(* IEC 61131-3 sources: teller/JD_Teller_LC2_V11/Network/HardwareNet, 1 file *)

(* ---- ONE_HardwareNet_Table.st ---- *)
#define OBJECTS_CONFIG

#include <.\lsl_st_can.h>
#include <.\lsl_st_hardwaretree.h>
//Define part of class HwBaseCDIAS
// Defines for Mutex Generation
#define CDIAS_STR_MUTEX_NAME_SEPERATOR ".."
#define CDIAS_MUTEX_NAME_END_LENGTH 5
#define CDIAS_MUTEX_NAME_MAX_LENGTH 32
//Define part of class CIO0xx
#define ID_CIO0xx 28

#define ID_CIO011 1
#define ID_CIO012 2
#define ID_CIO013 3
#define ID_CIO014 4
#define ID_CIO016 6
#define ID_CIO017 7

#define CIO0xx_Errormask 2#1111111110001111
//Define part of class Varan_Base
#ifndef _T_VARANBASE_H
#define _T_VARANBASE_H

#define	VARAN_PLL_OFFSET		16#0140
#define VARAN_MULTIPLE_OFFSET	16#01AC

// version of serial number validation (16#10 = 1.0)
#define SERNO_VALIDATION_VERSION 16#10

#define IsTransparent_IS_AVAILABLE

// Defines for Mutex Generation
#define VARAN_STR_MUTEX_NAME_SEPERATOR ".."
#define VARAN_MUTEX_NAME_END_LENGTH 5
#define VARAN_MUTEX_NAME_MAX_LENGTH 32

#endif // _T_VARANBASE_H
#include <.\lsl_st_pci.h>
#include "..\..\Class\DiasMasterMain\DiasMasterMain.h"
#include <.\lsl_st_kernel.h>
//Define part of class EEPROM
// Defines for Mutex Geeration
#define EEPROM_STR_MUTEX_NAME_SEPERATOR ".."
#define EEPROM_MUTEX_NAME_END_LENGTH 5
#define EEPROM_MUTEX_NAME_MAX_LENGTH 32
#include "..\..\Class\HwControl\HwControl.h"
//Define part of class SafetyManager
#define LogBufferSize 1000
#include "..\..\Class\SafetyManager\SafetyManager.h"
//Define part of class Varan_Can
#define VARAN_CAN_OS_VERSION	16#1100 + 226
#define CANBUS_INVALID_VALUE	-2147483393			//16#800000FF
//Define part of class VaranManager
#define SIZE_PAYLOAD_FRAME_HEADER_DO      36  // Const because datasize is in the Payload DOs
#define SIZE_PAYLOAD_IRQ_FRAME_HEADER_DO  38  // Const because datasize is in the Payload DOs

#define VM_MAX_POST_INIT_MODULES  1000
#include "..\..\Class\VaranManager\VaranManager.h"

FUNCTION GLOBAL TAB ONE_HardwareNet
-1$UINT, 0$UINT,
0$UINT, 0$UINT,

46$UDINT,
TO_UDINT(529317953), "_CanLib", 1$UINT, 10$UINT, 0$UINT,
TO_UDINT(4078275645), "_SerLib", 1$UINT, 31$UINT, 0$UINT,
TO_UDINT(781409069), "_VaranCanLib", 1$UINT, 10$UINT, 1$UINT,
TO_UDINT(415874427), "_VaranCanLibOS", 1$UINT, 10$UINT, 1$UINT,
TO_UDINT(3827919523), "_VaranSerLibOS", 1$UINT, 20$UINT, 3$UINT,
TO_UDINT(3907636883), "CAICIOAInputChannel", 2$UINT, 20$UINT, 2$UINT,
TO_UDINT(2472734913), "CAIInputChannel", 2$UINT, 20$UINT, 0$UINT,
TO_UDINT(1046309609), "CDias2DataMover", 1$UINT, 50$UINT, 1$UINT,
TO_UDINT(706219532), "ChannelBaseData", 1$UINT, 0$UINT, 0$UINT,
TO_UDINT(3340137983), "ChannelBaseDataWriteOnly", 1$UINT, 0$UINT, 0$UINT,
TO_UDINT(454909577), "CIO011_IM", 2$UINT, 50$UINT, 1$UINT,
TO_UDINT(2636333112), "CIO0xx", 2$UINT, 40$UINT, 0$UINT,
TO_UDINT(3867554050), "CIOOutputChannel", 2$UINT, 20$UINT, 1$UINT,
TO_UDINT(495304727), "CIV521", 1$UINT, 61$UINT, 1$UINT,
TO_UDINT(2756859380), "CIV_Base", 2$UINT, 61$UINT, 0$UINT,
TO_UDINT(658675781), "DAIInputChnl", 2$UINT, 10$UINT, 0$UINT,
TO_UDINT(3820159437), "Dias2DataMover", 1$UINT, 50$UINT, 1$UINT,
TO_UDINT(2647887450), "DiasMaster", 2$UINT, 30$UINT, 0$UINT,
TO_UDINT(3069482179), "DiasMasterC", 1$UINT, 70$UINT, 0$UINT,
TO_UDINT(3792535737), "DiasMasterMain", 2$UINT, 10$UINT, 0$UINT,
TO_UDINT(3076475114), "DiasMasterPostScan", 1$UINT, 0$UINT, 1$UINT,
TO_UDINT(2784851678), "EEPROM", 1$UINT, 11$UINT, 1$UINT,
TO_UDINT(3238133653), "Hub_Base", 1$UINT, 20$UINT, 1$UINT,
TO_UDINT(1770276445), "Hub_Base_Root", 2$UINT, 10$UINT, 1$UINT,
TO_UDINT(1800499398), "HwBaseCDIAS", 2$UINT, 50$UINT, 0$UINT,
TO_UDINT(2471641665), "HwControl", 3$UINT, 0$UINT, 1$UINT,
TO_UDINT(1193052171), "HwControlBase", 1$UINT, 10$UINT, 0$UINT,
TO_UDINT(4260294091), "HWRtPostScan", 1$UINT, 0$UINT, 1$UINT,
TO_UDINT(2326720416), "I2CCDIAS", 1$UINT, 6$UINT, 1$UINT,
TO_UDINT(3953068548), "JD_OR_Teller", 1$UINT, 0$UINT, 1$UINT,
TO_UDINT(2225119864), "MerkerEx", 1$UINT, 18$UINT, 4$UINT,
TO_UDINT(4209775899), "Pulser", 1$UINT, 1$UINT, 1$UINT,
TO_UDINT(3591333481), "RamFile", 1$UINT, 8$UINT, 1$UINT,
TO_UDINT(1799751072), "SafetyManager", 1$UINT, 42$UINT, 1$UINT,
TO_UDINT(1850111279), "String", 1$UINT, 10$UINT, 4$UINT,
TO_UDINT(2898603620), "StringInternal", 1$UINT, 70$UINT, 0$UINT,
TO_UDINT(4187542331), "SyncCall", 1$UINT, 20$UINT, 1$UINT,
TO_UDINT(862125188), "Varan_Base", 2$UINT, 2$UINT, 0$UINT,
TO_UDINT(206510048), "Varan_Can", 1$UINT, 40$UINT, 1$UINT,
TO_UDINT(3752737333), "Varan_DataMover", 1$UINT, 50$UINT, 1$UINT,
TO_UDINT(2940693151), "VaranManager", 2$UINT, 12$UINT, 0$UINT,
TO_UDINT(1989862026), "VaranManager_1", 1$UINT, 43$UINT, 1$UINT,
TO_UDINT(4035182347), "VaranManager_Base", 1$UINT, 20$UINT, 0$UINT,
TO_UDINT(803224590), "VaranManagerPostScan", 1$UINT, 1$UINT, 1$UINT,
TO_UDINT(3232495061), "VirtualBaseInit", 1$UINT, 3$UINT, 0$UINT,
TO_UDINT(1573657038), "WatchdogDias", 2$UINT, 10$UINT, 1$UINT,

1$UINT, TO_UDINT(2726984929), "CIV5211\_VARANCANLIB",

1$UINT, TO_UDINT(3666615371), "CIV5211\_VARANCANLIBOS",

1$UINT, TO_UDINT(2650501396), "CIV5211\_VARANSERLIBOS0",
1$UINT, TO_UDINT(3942400386), "CIV5211\_VARANSERLIBOS1",
1$UINT, TO_UDINT(1945440312), "CIV5211\_VARANSERLIBOS2",

1$UINT, TO_UDINT(3874057698), "CIO011_IM1\CAICIOAINPUTCHANNEL0",
1$UINT, TO_UDINT(2448317812), "CIO011_IM1\CAICIOAINPUTCHANNEL1",

1$UINT, TO_UDINT(407248868), "CIV5211\CDIAS2DATAMOVER",

_NO_ATTR, TO_UDINT(396609901), "CIO011_IM1",

1$UINT, TO_UDINT(325438698), "CIO011_IM1\CIOOUTPUTCHANNEL0",

_NO_ATTR, TO_UDINT(1241008), "CIV5211",

1$UINT, TO_UDINT(569811197), "CIV5211\DIAS2DATAMOVER",

1$UINT, TO_UDINT(2796364169), "CIV5211\DIAS2DATAMOVER\_BASE\DIASMASTERPOSTSCAN",

1$UINT, TO_UDINT(330460277), "CIV5211\DIAS2DATAMOVER\_BASE\EEPROM",

1$UINT, TO_UDINT(2268287070), "CIV5211\HUB_BASE0",

1$UINT, TO_UDINT(1776428101), "VARANMANAGER_11\HUB_BASE_ROOT0",

_NO_ATTR, TO_UDINT(2190789875), "HWCONTROL1",

1$UINT, TO_UDINT(1673205898), "HWCONTROL1\HWRTPOSTSCAN",

1$UINT, TO_UDINT(977257911), "CIV5211\DIAS2DATAMOVER\_BASE\I2CCDIAS",

_NO_ATTR, TO_UDINT(2206833861), "JD_OR1",

1$UINT, TO_UDINT(858933024), "CIO011_IM1\_BASE\_BASE\SERIALNOSTR\MERKEREX0",
1$UINT, TO_UDINT(2644417201), "CIV5211\DIAS2DATAMOVER\_BASE\SYNCCALL\_BASE\SERIALNOSTR\MERKEREX0",
1$UINT, TO_UDINT(3052700284), "CIV5211\DIAS2DATAMOVER\_BASE\WATCHDOGDIAS0\_BASE\SERIALNOSTR\MERKEREX0",
1$UINT, TO_UDINT(2330668179), "CIV5211\_BASE\SERIALNOSTR\MERKEREX0",

_NO_ATTR, TO_UDINT(155437646), "PULSER1",

1$UINT, TO_UDINT(4247336844), "CIV5211\_BASE\SERNOBACKUP",

1$UINT, TO_UDINT(1778590035), "HWCONTROL1\SAFETYMANAGER",

1$UINT, TO_UDINT(2060113651), "CIO011_IM1\_BASE\_BASE\SERIALNOSTR",
1$UINT, TO_UDINT(2623421091), "CIV5211\DIAS2DATAMOVER\_BASE\SYNCCALL\_BASE\SERIALNOSTR",
1$UINT, TO_UDINT(2991369526), "CIV5211\DIAS2DATAMOVER\_BASE\WATCHDOGDIAS0\_BASE\SERIALNOSTR",
1$UINT, TO_UDINT(2961157748), "CIV5211\_BASE\SERIALNOSTR",

1$UINT, TO_UDINT(1225390380), "CIV5211\DIAS2DATAMOVER\_BASE\SYNCCALL",

1$UINT, TO_UDINT(4278451883), "CIV5211\VARAN_CAN",

1$UINT, TO_UDINT(4189409080), "CIV5211\VARAN_DATAMOVER",

_NO_ATTR, TO_UDINT(2395414379), "VARANMANAGER_11",

1$UINT, TO_UDINT(4241828209), "VARANMANAGER_11\_BASE\VARANMASTERPOSTSCAN",

1$UINT, TO_UDINT(2365686840), "CIV5211\DIAS2DATAMOVER\_BASE\WATCHDOGDIAS0",

//Internal connections
0$UDINT,
31$UDINT,
TO_UDINT(8), "SerialNoStr", TO_UDINT(27),
TO_UDINT(8), "CAICIOAInputChannel0", TO_UDINT(5),
TO_UDINT(8), "CAICIOAInputChannel1", TO_UDINT(6),
TO_UDINT(8), "CIOOutputChannel0", TO_UDINT(9),
TO_UDINT(10), "SerialNoStr", TO_UDINT(30),
TO_UDINT(10), "SerNoBackup", TO_UDINT(25),
TO_UDINT(10), "Varan_DataMover", TO_UDINT(33),
TO_UDINT(10), "CDias2DataMover", TO_UDINT(7),
TO_UDINT(10), "Dias2DataMover", TO_UDINT(11),
TO_UDINT(10), "Hub_Base0", TO_UDINT(14),
TO_UDINT(10), "Varan_Can", TO_UDINT(32),
TO_UDINT(10), "_VaranCanLib", TO_UDINT(0),
TO_UDINT(10), "_VaranCanLibOS", TO_UDINT(1),
TO_UDINT(10), "_VaranSerLibOS0", TO_UDINT(2),
TO_UDINT(10), "_VaranSerLibOS1", TO_UDINT(3),
TO_UDINT(10), "_VaranSerLibOS2", TO_UDINT(4),
TO_UDINT(11), "DiasMasterPostScan", TO_UDINT(12),
TO_UDINT(11), "EEPROM", TO_UDINT(13),
TO_UDINT(11), "I2CCDIAS", TO_UDINT(18),
TO_UDINT(11), "WatchdogDias0", TO_UDINT(36),
TO_UDINT(11), "SyncCall", TO_UDINT(31),
TO_UDINT(16), "HWRtPostScan", TO_UDINT(17),
TO_UDINT(16), "SafetyManager", TO_UDINT(26),
TO_UDINT(27), "MerkerEx0", TO_UDINT(20),
TO_UDINT(28), "MerkerEx0", TO_UDINT(21),
TO_UDINT(29), "MerkerEx0", TO_UDINT(22),
TO_UDINT(30), "MerkerEx0", TO_UDINT(23),
TO_UDINT(31), "SerialNoStr", TO_UDINT(28),
TO_UDINT(34), "VaranMasterPostScan", TO_UDINT(35),
TO_UDINT(34), "Hub_Base_Root0", TO_UDINT(15),
TO_UDINT(36), "SerialNoStr", TO_UDINT(29),
0$UDINT,
33$UDINT,
TO_UDINT(0), "To_Varan_Can", TO_UDINT(32), "State",
TO_UDINT(1), "VaranIn", TO_UDINT(10), "State",
TO_UDINT(2), "VaranIn", TO_UDINT(10), "State",
TO_UDINT(3), "VaranIn", TO_UDINT(10), "State",
TO_UDINT(4), "VaranIn", TO_UDINT(10), "State",
TO_UDINT(5), "connectc", TO_UDINT(8), "State",
TO_UDINT(6), "connectc", TO_UDINT(8), "State",
TO_UDINT(7), "VaranIn", TO_UDINT(10), "State",
TO_UDINT(7), "To_DataMover", TO_UDINT(33), "State",
TO_UDINT(8), "MasterConnect", TO_UDINT(7), "Control",
TO_UDINT(9), "Connect", TO_UDINT(8), "State",
TO_UDINT(10), "VaranIn", TO_UDINT(15), "Control",
TO_UDINT(11), "SyncCall", TO_UDINT(31), "State",
TO_UDINT(11), "VaranIn", TO_UDINT(10), "State",
TO_UDINT(11), "To_DataMover", TO_UDINT(33), "State",
TO_UDINT(12), "MasterConnect", TO_UDINT(11), "Control",
TO_UDINT(13), "MasterConnect", TO_UDINT(11), "Control",
TO_UDINT(14), "VaranIn", TO_UDINT(10), "State",
TO_UDINT(15), "VaranConnect", TO_UDINT(34), "Control",
TO_UDINT(17), "toHwControlBase", TO_UDINT(16), "Control",
TO_UDINT(18), "MasterConnect", TO_UDINT(11), "Control",
TO_UDINT(19), "Out", TO_UDINT(8), "Output6",
TO_UDINT(26), "To_HwControl", TO_UDINT(16), "Control",
TO_UDINT(27), "DataBuffer", TO_UDINT(20), "m_udLength",
TO_UDINT(28), "DataBuffer", TO_UDINT(21), "m_udLength",
TO_UDINT(29), "DataBuffer", TO_UDINT(22), "m_udLength",
TO_UDINT(30), "DataBuffer", TO_UDINT(23), "m_udLength",
TO_UDINT(31), "MasterConnect", TO_UDINT(11), "Control",
TO_UDINT(32), "To_Varan_Base", TO_UDINT(10), "State",
TO_UDINT(33), "VaranIn", TO_UDINT(10), "State",
TO_UDINT(34), "To_HwControl", TO_UDINT(16), "Control",
TO_UDINT(35), "ManagerConnect", TO_UDINT(34), "Control",
TO_UDINT(36), "MasterConnect", TO_UDINT(11), "Control",

//Initialization values
0$UDINT,
70$UDINT,
TO_UDINT(1), "Index", TO_UDINT(0),//|HardwareNet.CIV5211\_VaranCanLibOS.Index;
TO_UDINT(2), "Index", TO_UDINT(0),//|HardwareNet.CIV5211\_VaranSerLibOS0.Index;
TO_UDINT(3), "Index", TO_UDINT(1),//|HardwareNet.CIV5211\_VaranSerLibOS1.Index;
TO_UDINT(4), "Index", TO_UDINT(2),//|HardwareNet.CIV5211\_VaranSerLibOS2.Index;
TO_UDINT(5), "channel", TO_UDINT(0),//|HardwareNet.CIO011_IM1\CAICIOAInputChannel0.channel;
TO_UDINT(5), "CyRt", TO_UDINT(1),//|HardwareNet.CIO011_IM1\CAICIOAInputChannel0.CyRt;
TO_UDINT(5), "CScale", TO_UDINT(10000),//|HardwareNet.CIO011_IM1\CAICIOAInputChannel0.CScale;
TO_UDINT(5), "BitResolution", TO_UDINT(12),//|HardwareNet.CIO011_IM1\CAICIOAInputChannel0.BitResolution;
TO_UDINT(5), "Neg", TO_UDINT(0),//|HardwareNet.CIO011_IM1\CAICIOAInputChannel0.Neg;
TO_UDINT(5), "EEOffset", TO_UDINT(16#48),//|HardwareNet.CIO011_IM1\CAICIOAInputChannel0.EEOffset;
TO_UDINT(6), "channel", TO_UDINT(1),//|HardwareNet.CIO011_IM1\CAICIOAInputChannel1.channel;
TO_UDINT(6), "CyRt", TO_UDINT(1),//|HardwareNet.CIO011_IM1\CAICIOAInputChannel1.CyRt;
TO_UDINT(6), "CScale", TO_UDINT(10000),//|HardwareNet.CIO011_IM1\CAICIOAInputChannel1.CScale;
TO_UDINT(6), "BitResolution", TO_UDINT(12),//|HardwareNet.CIO011_IM1\CAICIOAInputChannel1.BitResolution;
TO_UDINT(6), "Neg", TO_UDINT(0),//|HardwareNet.CIO011_IM1\CAICIOAInputChannel1.Neg;
TO_UDINT(6), "EEOffset", TO_UDINT(16#48),//|HardwareNet.CIO011_IM1\CAICIOAInputChannel1.EEOffset;
TO_UDINT(7), "CDIAS_BusAddress", TO_UDINT(0),//|HardwareNet.CIV5211\CDias2DataMover.CDIAS_BusAddress;
TO_UDINT(7), "MoverActive", TO_UDINT(1),//|HardwareNet.CIV5211\CDias2DataMover.MoverActive;
TO_UDINT(8), "Place", TO_UDINT(0),//|HardwareNet.CIO011_IM1.Place;
TO_UDINT(8), "Required", TO_UDINT(0),//|HardwareNet.CIO011_IM1.Required;
TO_UDINT(8), "RtCyInputs", TO_UDINT(1),//|HardwareNet.CIO011_IM1.RtCyInputs;
TO_UDINT(8), "RtCyOutputs", TO_UDINT(1),//|HardwareNet.CIO011_IM1.RtCyOutputs;
TO_UDINT(8), "Input3IRQMode", TO_UDINT(0),//|HardwareNet.CIO011_IM1.Input3IRQMode;
TO_UDINT(8), "CounterMode1and2", TO_UDINT(3),//|HardwareNet.CIO011_IM1.CounterMode1and2;
TO_UDINT(8), "AI_RtCy", TO_UDINT(1),//|HardwareNet.CIO011_IM1.AI_RtCy;
TO_UDINT(8), "AI1_CScale", TO_UDINT(10000),//|HardwareNet.CIO011_IM1.AI1_CScale;
TO_UDINT(8), "AI2_CScale", TO_UDINT(10000),//|HardwareNet.CIO011_IM1.AI2_CScale;
TO_UDINT(8), "AO_RtCy", TO_UDINT(1),//|HardwareNet.CIO011_IM1.AO_RtCy;
TO_UDINT(8), "AO_CScale", TO_UDINT(10000),//|HardwareNet.CIO011_IM1.AO_CScale;
TO_UDINT(9), "CScale", TO_UDINT(10000),//|HardwareNet.CIO011_IM1\CIOOutputChannel0.CScale;
TO_UDINT(10), "Required", TO_UDINT(0),//|HardwareNet.CIV5211.Required;
TO_UDINT(10), "Transparent", TO_UDINT(0),//|HardwareNet.CIV5211.Transparent;
TO_UDINT(10), "TimeBase", TO_UDINT(0),//|HardwareNet.CIV5211.TimeBase;
TO_UDINT(10), "TimeBaseOffset", TO_UDINT(0),//|HardwareNet.CIV5211.TimeBaseOffset;
TO_UDINT(10), "MoverActive", TO_UDINT(1),//|HardwareNet.CIV5211.MoverActive;
TO_UDINT(11), "DIAS_BusAddress", TO_UDINT(16#10000),//|HardwareNet.CIV5211\Dias2DataMover.DIAS_BusAddress;
TO_UDINT(14), "Splitter_Place", TO_UDINT(0),//|HardwareNet.CIV5211\Hub_Base0.Splitter_Place;
TO_UDINT(15), "Splitter_Place", TO_UDINT(0),//|HardwareNet.VaranManager_11\Hub_Base_Root0.Splitter_Place;
TO_UDINT(20), "ThreadSafe", TO_UDINT(0),//|HardwareNet.SerialNoStr\_base\_base\CIO011_IM1\MerkerEx0.ThreadSafe;
TO_UDINT(21), "ThreadSafe", TO_UDINT(0),//|HardwareNet.SerialNoStr\_base\SyncCall\_base\Dias2DataMover\CIV5211\MerkerEx0.ThreadSafe;
TO_UDINT(22), "ThreadSafe", TO_UDINT(0),//|HardwareNet.SerialNoStr\_base\WatchdogDias0\_base\Dias2DataMover\CIV5211\MerkerEx0.ThreadSafe;
TO_UDINT(23), "ThreadSafe", TO_UDINT(0),//|HardwareNet.SerialNoStr\_base\CIV5211\MerkerEx0.ThreadSafe;
TO_UDINT(24), "ResetIn", TO_UDINT(0),//|HardwareNet.Pulser1.ResetIn;
TO_UDINT(24), "ResetOut", TO_UDINT(0),//|HardwareNet.Pulser1.ResetOut;
TO_UDINT(25), "Setup", TO_UDINT(2#1101),//|HardwareNet._base\CIV5211\SerNoBackup.Setup;
TO_UDINT(27), "SingleRealloc", TO_UDINT(1),//|HardwareNet._base\_base\CIO011_IM1\SerialNoStr.SingleRealloc;
TO_UDINT(28), "SingleRealloc", TO_UDINT(1),//|HardwareNet._base\SyncCall\_base\Dias2DataMover\CIV5211\SerialNoStr.SingleRealloc;
TO_UDINT(29), "SingleRealloc", TO_UDINT(1),//|HardwareNet._base\WatchdogDias0\_base\Dias2DataMover\CIV5211\SerialNoStr.SingleRealloc;
TO_UDINT(30), "SingleRealloc", TO_UDINT(1),//|HardwareNet._base\CIV5211\SerialNoStr.SingleRealloc;
TO_UDINT(31), "Place", TO_UDINT(0),//|HardwareNet._base\Dias2DataMover\CIV5211\SyncCall.Place;
TO_UDINT(31), "Required", TO_UDINT(1),//|HardwareNet._base\Dias2DataMover\CIV5211\SyncCall.Required;
TO_UDINT(31), "TimeBase", TO_UDINT(0),//|HardwareNet._base\Dias2DataMover\CIV5211\SyncCall.TimeBase;
TO_UDINT(31), "TimeBaseOffset", TO_UDINT(0),//|HardwareNet._base\Dias2DataMover\CIV5211\SyncCall.TimeBaseOffset;
TO_UDINT(32), "Can_AddressOffset", TO_UDINT(16#4000),//|HardwareNet.CIV5211\Varan_Can.Can_AddressOffset;
TO_UDINT(32), "Index", TO_UDINT(0),//|HardwareNet.CIV5211\Varan_Can.Index;
TO_UDINT(33), "DPRAM_StartAddress", TO_UDINT(16#2000),//|HardwareNet.CIV5211\Varan_DataMover.DPRAM_StartAddress;
TO_UDINT(33), "DPRAM_StartAddress_SUBBus", TO_UDINT(16#2000),//|HardwareNet.CIV5211\Varan_DataMover.DPRAM_StartAddress_SUBBus;
TO_UDINT(33), "DPRAM_Size", TO_UDINT(4096),//|HardwareNet.CIV5211\Varan_DataMover.DPRAM_Size;
TO_UDINT(33), "CodeStartAddress", TO_UDINT(16#8000),//|HardwareNet.CIV5211\Varan_DataMover.CodeStartAddress;
TO_UDINT(33), "CodeSize", TO_UDINT(4096),//|HardwareNet.CIV5211\Varan_DataMover.CodeSize;
TO_UDINT(33), "TimeSliceErrorOn", TO_UDINT(1),//|HardwareNet.CIV5211\Varan_DataMover.TimeSliceErrorOn;
TO_UDINT(34), "VaranManagerTime", TO_UDINT(1000000),//|HardwareNet.VaranManager_11.VaranManagerTime;
TO_UDINT(34), "VaranManagerNr", TO_UDINT(0),//|HardwareNet.VaranManager_11.VaranManagerNr;
TO_UDINT(34), "PayloadFrame", TO_UDINT(0),//|HardwareNet.VaranManager_11.PayloadFrame;
TO_UDINT(34), "PayloadMEMWrite", TO_UDINT(0),//|HardwareNet.VaranManager_11.PayloadMEMWrite;
TO_UDINT(34), "PayloadMEMRead", TO_UDINT(0),//|HardwareNet.VaranManager_11.PayloadMEMRead;
TO_UDINT(36), "Place", TO_UDINT(0),//|HardwareNet._base\Dias2DataMover\CIV5211\WatchdogDias0.Place;
TO_UDINT(36), "Required", TO_UDINT(1),//|HardwareNet._base\Dias2DataMover\CIV5211\WatchdogDias0.Required;
TO_UDINT(36), "TimeBase", TO_UDINT(0),//|HardwareNet._base\Dias2DataMover\CIV5211\WatchdogDias0.TimeBase;
TO_UDINT(36), "TimeBaseOffset", TO_UDINT(0),//|HardwareNet._base\Dias2DataMover\CIV5211\WatchdogDias0.TimeBaseOffset;

//Symbolic initialization values
0$UDINT,
0$UDINT,

//Initialization of string values
0$UDINT,
0$UDINT,

//Configuration of tasks (RealTime, Cyclic, Background)
0$UDINT,
2$UDINT,
TO_UDINT(16), (1)$UDINT, 0$DINT, 	//HWCONTROL1
TO_UDINT(17), (1)$UDINT, 4194304$DINT, 	//HWCONTROL1\HWRTPOSTSCAN

0$UDINT,
2$UDINT,
TO_UDINT(24), (100)$UDINT, 4194303$DINT, 	//PULSER1
TO_UDINT(16), (1)$UDINT, 8388607$DINT, 	//HWCONTROL1

0$UDINT,
0$UDINT,

//External connections
0$UDINT,
0$UDINT,

//Magic internal connections
0$UDINT,
18$UDINT,
TO_UDINT(5), "TypeofChannel", TO_UDINT(8), "AI1_TypeofChannel",
TO_UDINT(5), "CyRt", TO_UDINT(8), "AI_RtCy",
TO_UDINT(5), "CScale", TO_UDINT(8), "AI1_CScale",
TO_UDINT(5), "CBias", TO_UDINT(8), "AI1_CBias",
TO_UDINT(5), "CInvert", TO_UDINT(8), "AI1_CInvert",
TO_UDINT(6), "TypeofChannel", TO_UDINT(8), "AI2_TypeofChannel",
TO_UDINT(6), "CyRt", TO_UDINT(8), "AI_RtCy",
TO_UDINT(6), "CScale", TO_UDINT(8), "AI2_CScale",
TO_UDINT(6), "CBias", TO_UDINT(8), "AI2_CBias",
TO_UDINT(6), "CInvert", TO_UDINT(8), "AI2_CInvert",
TO_UDINT(7), "MoverActive", TO_UDINT(10), "MoverActive",
TO_UDINT(9), "CScale", TO_UDINT(8), "AO_CScale",
TO_UDINT(9), "CBias", TO_UDINT(8), "AO_CBias",
TO_UDINT(9), "CInvert", TO_UDINT(8), "AO_CInvert",
TO_UDINT(26), "SafetyDomainTimeout", TO_UDINT(16), "SafetyDomainTimeout",
TO_UDINT(32), "Pll_Prescaler", TO_UDINT(10), "Pll_Prescaler",
TO_UDINT(32), "CallUserRt", TO_UDINT(10), "CallUserRt",
TO_UDINT(32), "ISOCanOn", TO_UDINT(10), "ISOCanOn",

//Configuration of timeslots of tasks (RealTime, Cyclic)
#ifdef __LSLLDR_TIMESLOTS__
0$UDINT,
0$UDINT,

0$UDINT,
0$UDINT,

#endif //__LSLLDR_TIMESLOTS__

//MultiMaster connections
#ifdef __LSLLDR_MULTIMASTER__
0$UDINT,
0$UDINT,
#endif //__LSLLDR_MULTIMASTER__

END_FUNCTION
